FUNCTION_BLOCK FB_Einlauf
VAR_INPUT
END_VAR
VAR_OUTPUT
END_VAR
VAR
END_VAR

IF GVL_IO.xLichtschranke_Einlauf AND GVL_IO.xServo_Einlauf_GS THEN
    GVL_IO.xEinlaufBereit := TRUE;
ELSIF NOT GVL_IO.xLichtschranke_Einlauf THEN
    GVL_IO.xEinlaufBereit := FALSE;
END_IF

END_FUNCTION_BLOCK

(* stored: Version 1.1.0.1
   POU FB_Einlauf: Id {1fbece50-0130-45db-9784-d8a45e6787fd}, SpecialFunc None *)
